//			Left				Visibility 5x / Error/select				right
//	 ___________________________________________________________________________________
//	|				| l |                                            |r |				|
//	|               | e |      headerText :  addText                 |i |               |
//	|  	 /          | f |--------------------------------------------|g |          \   	|
//	|	/           | t |    infoText1   		|	infoText2		 |ht|           \  	|		
//  |	\           | . |                       |                    |. |           /   |
//  | 	 \          | st|--------------------------------------------|st|          /    |
// 	| Left.key.text	| at|    infoText3          |	infoText4        |at| right.key.text|
//	|_______________|_us|_______________________|____________________|us|_______________|

// sort  [1 - n] änder die Anzeige Reihenfolge

END_FUNCTION_BLOCK

// DUTs/HMI_ManualFnc/FB_ManualFncFull
{attribute 'OPC.UA.DA' := '1'}
FUNCTION_BLOCK FB_ManualFncFull EXTENDS FB_ManualFncBody
VAR_INPUT
	left					:	FB_ManualFncKey;
	right					:	FB_ManualFncKey;
END_VAR

//			Left				Visibility 5x / Error/select				right
//	 ___________________________________________________________________________________
//	|				| l |                                            |r |				|
//	|               | e |      headerText :  addText                 |i |               |
//	|  	 /          | f |--------------------------------------------|g |          \   	|
//	|	/           | t |    infoText1   		|	infoText2		 |ht|           \  	|		
//  |	\           | . |                       |                    |. |           /   |
//  | 	 \          | st|--------------------------------------------|st|          /    |
// 	| Left.key.text	| at|    infoText3          |	infoText4        |at| right.key.text|
//	|_______________|_us|_______________________|____________________|us|_______________|

// sort  [1 - n] änder die Anzeige Reihenfolge

END_FUNCTION_BLOCK

// DUTs/HMI_ManualFnc/FB_ManualFncKey
{attribute 'OPC.UA.DA' := '1'}
FUNCTION_BLOCK FB_ManualFncKey
VAR_INPUT
	key					:	FB_ManualFncKeyBasic;
	status				:	FB_ManualFncStatus;
END_VAR

END_FUNCTION_BLOCK

// DUTs/HMI_ManualFnc/FB_ManualFncKeyBasic
{attribute 'OPC.UA.DA' := '1'}
FUNCTION_BLOCK FB_ManualFncKeyBasic
VAR_INPUT
	text				:	STRING;
	cssAttribut			: 	STRING;
	disable				:	BOOL;
	userLevel			:	INT;
	liveBit				:	BOOL;
	q					:	BOOL;
	colorChange			:	BOOL := FALSE;
	hide				:	ST_KeyHide;	
END_VAR

END_FUNCTION_BLOCK

// DUTs/HMI_ManualFnc/FB_ManualFncStatus
{attribute 'OPC.UA.DA' := '1'}
FUNCTION_BLOCK FB_ManualFncStatus
VAR_INPUT
	text				:	STRING;
	colorChange			:	BOOL := FALSE;
	hide				:	ST_StatusHide;	
END_VAR

END_FUNCTION_BLOCK
